{attribute 'qualified_only'}
VAR_GLOBAL CONSTANT
	nZONES_MAX_NO			:UINT := 4;			(* Amount of control zones *)
END_VAR

(* stored: Version 1.1.0.1, ProductVersion 3.1.4024.15
   GVL GVL_GFX4IR: Id {4cf04c45-faaf-4b4d-94de-7f1c43babdcb} *)
